// TIA Portal V18 export
VAR_GLOBAL   // PLC tag table "Setup"
   Tag_19 AT %I0.0 : Bool;
END_VAR
VAR_GLOBAL CONSTANT   // user constants
   ModeZone_Setup_Const : Int := 12;
   Station_Setup_Const : Int := 20;
   Position_Setup_Const : Int := 1;
   Equipment_Setup_Const : Int := 10;
   ThisProcess : Int := 1;
   ThisWorkshop : Int := 1;
   Connection_Setup_Const : Int := 30;
   ContractID_Setup_Const : Int := 24;
   ITConnectionName : String := 'PLC_AREA_01';
   Parameter_Setup_Const : Int := 20;
   WorkPlace_Setup_Const : Int := 16;
   Total_User_Const : Int := 200;
   User_Roles_Const : Int := 100;
   ProductionSequenceList_Setup_Const : Int := 30;   // Quantidade de produtos que podemos ter por posto
   listTypeReason_Const : Int := 200;
   ITConnectionID : Word := W#16#101;
   Signal_Setup_Const : Int := 8;
   ShiftList_Setup_Const : Int := 3;
   Quantidade_task : Int := 10;
   Tamanho_POPID : Int := 7;
   nProcess : Int := 1;
   Quantidade_Paradas_Matriz : Int := 2;
END_VAR
